// Fire-and-forget message whose severity and text come from the event catalog.
FUNCTION_BLOCK FB_CatalogMessage EXTENDS FB_CatalogEventBase IMPLEMENTS I_Message
VAR
	_fbMessage	: FB_TcMessage;
END_VAR

METHOD PROTECTED CreateEvent : HRESULT
VAR_INPUT
	stEventEntry	: TcEventEntry;
	ipSourceInfo	: I_TcSourceInfo;
END_VAR
CreateEvent := _fbMessage.CreateEx(stEventEntry := stEventEntry, ipSourceInfo := ipSourceInfo);
END_METHOD

METHOD Send : HRESULT
VAR
	sText	: T_MaxString;
END_VAR
IF NOT EnsureCreated() THEN
	Send := _hrLast;
	RETURN;
END_IF

sText := BuildText();
_fbMessage.ipArguments.Clear().AddString(sText);
_hrLast := _fbMessage.Send(0);
Send := _hrLast;
END_METHOD

END_FUNCTION_BLOCK

(* stored: Version 1.1.0.1, ProductVersion 3.1.4026.26
   POU FB_CatalogMessage: Id {9385f519-9b28-4e74-9657-543aaa1eddd9}, SpecialFunc None
   Method CreateEvent: Id {8bbcde68-6510-4aef-a360-593251362ffa}
   Method Send: Id {2bf7a438-844d-4c87-a04e-c16c87ceb717} *)
